PROGRAM PRG_Wash
VAR
    bStart : BOOL;
    bMoto : BOOL;
    bAuto : BOOL;
    nStep : INT;
END_VAR

nStep := nStep + 1;

TRANSITION T_Bare:
bStart AND NOT bAuto
END_TRANSITION

TRANSITION T_Semicolon:
(bMoto OR bAuto) AND nStep = 1;
END_TRANSITION

TRANSITION T_Name:
bStart;
END_TRANSITION

TRANSITION T_Comment:
nStep > 2; // after the second step
END_TRANSITION

TRANSITION T_Assign:
T_Assign := bMoto AND bStart;
END_TRANSITION

END_PROGRAM

(* stored: Version 1.1.0.1, ProductVersion 3.1.4024.12
   POU PRG_Wash: Id {00000000-0000-0000-0000-000000000101}, SpecialFunc None
   Transition T_Bare: Id {00000000-0000-0000-0000-000000000102}
   Transition T_Semicolon: Id {00000000-0000-0000-0000-000000000103}
   Transition T_Name: Id {00000000-0000-0000-0000-000000000104}
   Transition T_Comment: Id {00000000-0000-0000-0000-000000000105}
   Transition T_Assign: Id {00000000-0000-0000-0000-000000000106} *)
